FUNCTION F_CreateTurbineCMD
VAR_INPUT
// 	nID				: UDINT;
END_VAR
VAR_OUTPUT
	sTurbineCmd		: S_TURBINECMD;
END_VAR
VAR
	temp: SINT;
	nID: UDINT;
END_VAR


FOR nID := 1 TO c_nNumTurbines DO
	temp := fbWTURBINE[nID].WTURBINELD0.WTUR1.TurOp.st_.stVal.iAny;
	sTurbineCmd.bEnable[nID] :=  SINT_TO_BOOL(temp);
	sTurbineCmd.bEmergencyStop[nID] := FALSE;
	sTurbineCmd.eCtrlMode[nID] := fbWTURBINE[nID].WTURBINELD0.WTUR1.TurCtl.st_.stVal.iAny;
	sTurbineCmd.fWSpt[nID] 	:= fbWTURBINE[nID].WTURBINELD0.WTUR1.DmdWSpt.val.mxVal.fValue;
	sTurbineCmd.fYawSpt[nID] := fbWTURBINE[nID].WTURBINELD0.WYAW1.YwAngSpt.val.mxVal.fValue;
END_FOR

END_FUNCTION

(* stored: Version 1.1.0.1
   POU F_CreateTurbineCMD: Id {8091cc33-872d-4ec0-b1d3-c128684dee94}, SpecialFunc None *)
